(*
SPDX-FileCopyrightText: © 2026 Oleksandr Tiutyk <trofimich@gmail.com>
SPDX-License-Identifier: MIT
License: https://opensource.org/license/mit
*)

(*!
<summary>
Beckhoff bidirectional counter channel process image.
</summary>
<description>
Aggregates input status/value (COUNTER_INPUT_CHANNEL) and output control/preset (COUNTER_OUTPUT_CHANNEL) for
one counter channel.
When used for I/O, link located fields or their containing buffers to the matching selected PDOs.
The record is not a packed wire buffer; compiler padding is not part of the device specification.
Unlinked/default values do not prove valid I/O. The caller evaluates bus/channel validity before use.
Use one owner task per instance and externally synchronize other access; multi-field snapshots are not atomic.
Copies store data without creating hardware links. Keep borrowed field references valid while consumers are bound.
This passive record performs no validation, synchronization, configuration or protocol advancement.
</description>
*)
TYPE COUNTER_CHANNEL :
STRUCT
	In : COUNTER_INPUT_CHANNEL;
	Out : COUNTER_OUTPUT_CHANNEL;
END_STRUCT
END_TYPE

(* stored: Version 1.1.0.1, ProductVersion 3.1.4026.20
   DUT COUNTER_CHANNEL: Id {0a7b98e6-4535-4d12-b736-ec2b88ce0783} *)
